// TIA Portal V20 export
Screen "Pop-up_EUCHNER_MGB_LEGEND_Popup"  380x408
  ScreenItem "Background" at 0,0 size 380x408  Type=HmiRectangle
  ScreenItem "Textfeld_Legende" at 1,1 size 378x25  Type=HmiTextBox
  ScreenItem "Textfeld_1" at 10,153 size 155x20  Type=HmiTextBox
  ScreenItem "Textfeld_3" at 10,55 size 155x20  Type=HmiTextBox
  ScreenItem "Textfeld_4" at 10,87 size 155x20  Type=HmiTextBox
  ScreenItem "Textfeld_5" at 10,109 size 155x20  Type=HmiTextBox
  ScreenItem "Textfeld_6" at 10,131 size 155x20  Type=HmiTextBox
  ScreenItem "Textfeld_10" at 170,153 size 200x20  Type=HmiTextBox
  ScreenItem "Textfeld_11" at 170,45 size 200x40  Type=HmiTextBox
  ScreenItem "Textfeld_12" at 170,87 size 200x20  Type=HmiTextBox
  ScreenItem "Textfeld_13" at 170,109 size 200x20  Type=HmiTextBox
  ScreenItem "Textfeld_14" at 170,131 size 200x20  Type=HmiTextBox
  ScreenItem "Textfeld_15" at 10,178 size 100x20  Type=HmiTextBox
  ScreenItem "Textfeld_16" at 75,201 size 300x40  Type=HmiTextBox
  ScreenItem "Textfeld_17" at 75,243 size 300x20  Type=HmiTextBox
  ScreenItem "Textfeld_18" at 75,264 size 300x39  Type=HmiTextBox
  ScreenItem "Textfeld_19" at 75,345 size 300x20  Type=HmiTextBox
  ScreenItem "Textfeld_20" at 75,366 size 300x39  Type=HmiTextBox
  ScreenItem "Cancel Mode" at 289,1 size 90x60  Type=HmiButton
  ScreenItem "Handle_Top_DoorOff" at 10,283 size 17x0  Type=HmiLine
  ScreenItem "Handle_Top_DoorOff_1" at 10,323 size 17x0  Type=HmiLine
  ScreenItem "Lock" at 10,345 size 16x16  Type=HmiGraphicView
  ScreenItem "Pushbutton_Left_ON" at 0,0 size 100x30  Type=HmiCircle
  ScreenItem "Pushbutton_Right_ON" at 0,0 size 100x30  Type=HmiCircle
  ScreenItem "Line_Automatic" at 16,221 size 6x0  Type=HmiLine
  ScreenItem "Frame_Door" at 58,216 size 6x10  Type=HmiRectangle
  ScreenItem "Doorhandle" at 58,221 size 3x0  Type=HmiLine
  ScreenItem "Pushbutton_Middle_ON" at 0,0 size 100x30  Type=HmiCircle
  ScreenItem "Text_" at 36,214 size 8x14  Type=HmiTextBox
  ScreenItem "Textfeld_2" at 75,304 size 300x39  Type=HmiTextBox
  ScreenItem "Frame_Yellow_R25" at 0,0 size 100x30  Type=HmiCircle
  ScreenItem "Switch_Shadow_R6" at 0,0 size 100x30  Type=HmiCircle
  ScreenItem "Switch_Red_R6" at 0,0 size 100x30  Type=HmiCircle
  ScreenItem "Handle_Down_DoorClosed" at 10,243 size 6x22  Type=HmiRectangle
